(* IEC 61131-3 sources: 2026_Projet_YGO_ExcavatriceDragage/CODE_BACKUP/CODE_20260907_ChantierWeekEnd_v0.6.43/L_SIMULATION, 5 files *)

(* ---- FB_Sim_Encoder.st ---- *)
(* ═══════════════════════════════════════════════════════════════
   🧪 FB_Sim_Encoder — Simulation physique d'un codeur absolu de treuil
   ───────────────────────────────────────────────────────────────
   📄 Doc métier : DOC/AF/AF_Partie-13_Fonction_Simulation_v2.5.md
   🧩 Brique réduite (Partie3 §1bis, "briques E/S & diagnostics") : pas de contrat
      Enable/Reset/Error complet, pas de StartStop/SafeStop — outil de banc, pas
      du métier machine.
   🎯 Rôle : fait "compter" un codeur absolu comme si le treuil tournait
      réellement, à partir des relais de sens commandés et du palier de vitesse courant.
   📥 Enable      : simulation active (SimulationModeActive AND NOT BusEncoderMxIsReal)
   📥 RelayFwd/RelayRev : sens commandé (contacteurs de sens du treuil)
   📥 StepNumber  : palier vitesse courant (1..5) — ex. instWinchM1.StepNumber
      Vitesse = interpolation linéaire : palier 1 → MinSpeedMps (1 m/s), palier 5 → MaxSpeedMps (2 m/s).
   📥 PresetCmd   : TRUE le cycle où un preset (homing) doit être appliqué (PresettTrigCmd = 2)
   📥 PresetValue : valeur brute à charger lors du preset
   📥 SpeedScaleFactor : facteur fin de confort (réglable à chaud, sans recompiler). Défaut 1.0 = vitesse
      réelle telle que définie par MinSpeedMps/MaxSpeedMps/PointsPerRev/CableM_PerRev/CycleTimeS.
   📤 RawPosOut   : position brute simulée (UDINT), à aiguiller à la place de la valeur
      EtherCAT réelle quand le device n'est pas Operational (voir PRG_02_Encoders.st)
   `RawPos` en `VAR_IN_OUT`, référencé depuis `GVL_PERSISTENT`
      (même pattern que `Calib` dans `FB_Encoder_Homing`) — `PERSISTENT` n'est valide que sur du
      `VAR_GLOBAL` en CODESYS, pas sur une variable locale de FB. Un vrai codeur absolu physique
      conserve son comptage brut même à travers un reset FROID (indépendant de l'automate).
   ═══════════════════════════════════════════════════════════════ *)

// === DECLARATION (à coller dans la partie déclaration du POU FB_Sim_Encoder) ===

FUNCTION_BLOCK PUBLIC FB_Sim_Encoder
VAR_INPUT
    Enable           : BOOL;   (* --> [CMD] Active la simulation *)
    RelayFwd         : BOOL;   (* --> [HW] Sens commandé avant *)
    RelayRev         : BOOL;   (* --> [HW] Sens commandé arrière *)
    StepNumber       : INT;    (* --> [CMD] Palier vitesse courant (1..5, 0 = arrêt) *)
    PresetCmd        : BOOL;   (* --> [CMD] Applique un preset (homing) *)
    PresetValue      : UDINT;   (* --> [CFG] Valeur brute à charger au preset *)
    SpeedScaleFactor : REAL := 1.0;   (* --> [CFG] Facteur fin de confort (défaut 1.0) *)
    CoastDistanceM   : REAL := 0.0;   (* --> [CFG] Distance de roulis inertiel apres coupure des relais (m). 0 = arret net (defaut). >0 = le treuil continue a vitesse palier 1 dans le dernier sens sur CoastDistanceM metres -> modelise l'anticipation d'arret mecanique (ex. benne). *)
    PresetLatencyCycles : INT := 3;   (* --> [CFG] Nb cycles automate avant application du preset (referencement non instantane) *)
    TestOffsetCmd    : BOOL;          (* --> [TST] Front montant = applique TestOffsetPts (test banc) *)
    TestOffsetPts    : DINT := 0;     (* --> [TST] Décalage signé à appliquer (points bruts) *)
    // 📐 Paramètres physiques du treuil (mêmes valeurs que FB_Encoder_Scale) + vitesse réelle.
    // Vitesse simulée = interpolation linéaire du palier : palier 1 → MinSpeedMps, palier 5 → MaxSpeedMps.
    MinSpeedMps      : REAL := 1.0;    (* --> [CFG] Vitesse palier 1 (m/s) *)
    MaxSpeedMps      : REAL := 2.0;    (* --> [CFG] Vitesse palier 5 (m/s) *)
    PointsPerRev     : UDINT := 8192;  (* --> [CFG] Résolution codeur (pts/tour) *)
    CableM_PerRev    : REAL := 2.0;    (* --> [CFG] Développement câble (m/tour) *)
    CycleTimeS       : REAL := 0.010;  (* --> [CFG] Période tâche PLC (s) — MainTask 10 ms *)
END_VAR
VAR_OUTPUT
    RawPosOut   : UDINT;   (* <-- [DIAG] Position brute simulée *)
    RawSpdOut   : DINT;    (* <-- [DIAG] Vitesse brute simulée (0x6031:01 en 0.1 RPM) *)
END_VAR
VAR_IN_OUT
    RawPos      : UDINT;   (* <-> [BUS] Référence _SimEncoderRawPosM1/M2 (survit au reset froid) *)
END_VAR
VAR
    Increment      : UDINT;              (* . [LOC] Points ajoutés par cycle *)
    EffStep        : INT;               (* . [LOC] Pas borné (>= 1) *)
    SpeedMps       : REAL;              (* . [LOC] Vitesse simulée (m/s) *)
    TestOffsetEdge : R_TRIG;             (* . [LOC] Front TestOffsetCmd *)
    PresetEdge     : R_TRIG;             (* . [LOC] Front montant PresetCmd *)
    PresetPending  : BOOL;               (* . [LOC] Preset en attente d'application (latence) *)
    PresetCount    : INT;                (* . [LOC] Compteur cycles de latence restants *)
    IncrStep1      : UDINT;              (* . [LOC] Increment par cycle a vitesse palier 1 (pour le roulis) *)
    MovingDir      : INT;                (* . [LOC] Dernier sens actif : +1 avant, -1 arriere, 0 arret *)
    CoastPtsLeft   : REAL;               (* . [LOC] Roulis inertiel restant (points bruts) *)
END_VAR

// === IMPLEMENTATION (à coller dans le corps ST du POU FB_Sim_Encoder) ===

{region "§1 Gate"}
IF NOT Enable THEN
    RawPosOut := RawPos;
    RETURN;
END_IF;
{endregion}

{region "§2 Injection test"}
// Injection test banc : VRAI saut de position (comme un glissement réel),
// pour tester Concept 1 / Méca E ET le rattrapage joystick (voir GVL_Simulation bandeau).
TestOffsetEdge(CLK := TestOffsetCmd);
IF TestOffsetEdge.Q THEN
    RawPos := DINT_TO_UDINT(UDINT_TO_DINT(RawPos) + TestOffsetPts);
END_IF;
{endregion}

{region "§3 Comptage"}
// 🎚️ Vitesse simulée = interpolation linéaire du palier (palier 1 → MinSpeedMps, palier 5 → MaxSpeedMps),
// pas par pas de (Max−Min)/4. Palier 0 (arrêt) ramène au palier 1 mais aucun mouvement n'est
// appliqué tant que RelayFwd/RelayRev = FALSE (section plus bas).
EffStep  := MAX(StepNumber, 1);
SpeedMps := MinSpeedMps + (INT_TO_REAL(EffStep) - 1.0) * ((MaxSpeedMps - MinSpeedMps) / 4.0);
// Points par cycle = vitesse (m/s) × points par mètre × période tâche (s) × facteur confort.
Increment := REAL_TO_UDINT(SpeedMps * (UDINT_TO_REAL(PointsPerRev) / CableM_PerRev) * CycleTimeS * SpeedScaleFactor);
// Increment "lent" (palier 1) : vitesse du roulis inertiel apres coupure des relais.
IncrStep1 := REAL_TO_UDINT(MinSpeedMps * (UDINT_TO_REAL(PointsPerRev) / CableM_PerRev) * CycleTimeS * SpeedScaleFactor);

// Front du preset : lance la latence de referencement (le codeur réel n'est pas
// instantane — il met PresetLatencyCycles cycles a se re-referencer apres le front).
PresetEdge(CLK := PresetCmd);
IF PresetEdge.Q THEN
    PresetPending := TRUE;
    PresetCount := PresetLatencyCycles;
END_IF;

// Pendant l'attente, la position brute est conservee (le codeur n'a pas encore re-reference).
// Le mouvement est gelé pendant la latence, comme un codeur réel en cours de referencement.
IF PresetPending THEN
    IF PresetCount > 0 THEN
        PresetCount := PresetCount - 1;
    ELSE
        // Latence écoulée : applique la valeur cible du preset.
        RawPos := PresetValue;
        PresetPending := FALSE;
    END_IF;
ELSIF RelayFwd THEN
    RawPos := RawPos + Increment;
    MovingDir := 1;
    CoastPtsLeft := CoastDistanceM * (UDINT_TO_REAL(PointsPerRev) / CableM_PerRev);
ELSIF RelayRev THEN
    IF RawPos >= Increment THEN
        RawPos := RawPos - Increment;
    ELSE
        RawPos := 0;
    END_IF;
    MovingDir := -1;
    CoastPtsLeft := CoastDistanceM * (UDINT_TO_REAL(PointsPerRev) / CableM_PerRev);
ELSE
    // Relais coupes : roulis inertiel (anticipation d'arret mecanique). Le treuil
    // continue a vitesse palier 1 dans le dernier sens jusqu'a epuisement de CoastPtsLeft.
    IF (CoastPtsLeft >= 1.0) AND (MovingDir <> 0) THEN
        IF MovingDir = 1 THEN
            RawPos := RawPos + IncrStep1;
        ELSIF RawPos >= IncrStep1 THEN
            RawPos := RawPos - IncrStep1;
        ELSE
            RawPos := 0;
        END_IF;
        CoastPtsLeft := CoastPtsLeft - UDINT_TO_REAL(IncrStep1);
    ELSE
        MovingDir := 0;
        CoastPtsLeft := 0.0;
    END_IF;
END_IF;
{endregion}

{region "§4 Sortie"}
RawPosOut := RawPos;
// Formule inverse vitesse brute EtherCAT CoE (0.1 RPM) :
// SpdValue = (V_mps * 60.0) / (0.1 * CableM_PerRev) = V_mps * 300.0 (sur tambour 2m)
IF (MovingDir <> 0) AND (CableM_PerRev > 0.0) THEN
    IF MovingDir = 1 THEN
        RawSpdOut := REAL_TO_DINT((SpeedMps * 60.0) / (0.1 * CableM_PerRev) * SpeedScaleFactor);
    ELSE
        RawSpdOut := -REAL_TO_DINT((SpeedMps * 60.0) / (0.1 * CableM_PerRev) * SpeedScaleFactor);
    END_IF;
ELSE
    RawSpdOut := 0;
END_IF;
{endregion}

END_FUNCTION_BLOCK

(* ---- FB_Sim_Joystick.st ---- *)
(* ═══════════════════════════════════════════════════════════════
   🧪 FB_Sim_Joystick — Simulation des entrées brutes joystick (bus CAN hors ligne)
   ───────────────────────────────────────────────────────────────
   📄 Doc métier : DOC/AF/AF_Partie-13_Fonction_Simulation_v2.5.md
   🧩 Brique réduite (Partie3 §1bis) : outil de banc, pas du métier machine.
   🎯 Rôle : remplace l'ancien bypass homme-mort codé en dur dans `FB_Joystick`
      (`GVL_DEBUG.DBG_DeadmanBypass_TEST`, qui forçait `DeadmanArmed` en
      permanence — un vrai contournement de sécurité). Ici, on simule les
      ENTRÉES BRUTES du capteur (`RawX`/`RawY`/`RawButton`) : le homme-mort réel
      de `FB_Joystick` reste pleinement actif et doit toujours être "actionné"
      (forcer `RawButton` en instance CODESYS) pour armer — comportement
      métier testé pour de vrai, pas contourné.
   🕹️ Comportement dynamique (conception validée) :
      - Ascending : bouton actif → `RawX`/`RawY` monte de `NeutralRaw` vers la cible
        (0 ou `MaxRaw`) en `RiseTimeS`, avec un bruit pseudo-aléatoire léger.
      - Dépassement (`OvershootActive`) : la cible de montée DÉPASSE la butée
        (MaxRaw+AMT ou 0−AMT) → déclenche le défaut capteur hors plage.
      - Retombée : bouton relâché → descente LINÉAIRE en `FallTimeMs` vers le neutre.
      - Bagotement (`BagotementActive`) : au retour, petit balancement de quelques %
        autour du neutre avant de se stabiliser.
   📥 Enable        : simulation active (SimulationModeActive AND NOT BusJoystickSignalIsReal)
   📥 NeutralRaw    : valeur brute simulée au repos (voir GVL_Simulation.TstJoystickForceNeutralRaw)
   📥 MaxRaw        : valeur brute simulée à fond (voir GVL_Simulation.TstJoystickForceMaxRaw)
   📥 Btn*          : boutons directionnels (1 seul impose une butée d'axe ; 0 ou ≥2 = neutre)
   📥 OvershootActive : bagotement au retour (test mouvement parasite)
   📥 RiseTimeS / FallTimeMs / CycleTimeS : dynamique temporelle (pattern FB_Sim_Encoder)
   📤 RawX/RawY     : valeurs brutes dynamiques (neutre = NeutralRaw)
   📤 RawButton     : homme-mort brut = un bouton directionnel actif
   💡 Note d'application : en vue instance CODESYS, forcer `RawX`/`RawY` à `MaxRaw` (ou une
      valeur intermédiaire) pour simuler un débattement, et `RawButton` à `TRUE` pour simuler
      l'appui homme-mort — exactement comme on forcerait le vrai capteur.
   ═══════════════════════════════════════════════════════════════ *)

// === DECLARATION (à coller dans la partie déclaration du POU FB_Sim_Joystick) ===

FUNCTION_BLOCK PUBLIC FB_Sim_Joystick
VAR_INPUT
    Enable              : BOOL;   (* --> [CMD] Active la simulation *)
    NeutralRaw          : INT := 5000;   (* --> [CFG] Valeur brute au repos (neutre) *)
    MaxRaw              : INT := 10000;   (* --> [CFG] Valeur brute à fond *)
    BtnLeft_Rev_TREMIE  : BOOL;   (* --> [TST] Bouton gauche : X→0, Y→neutre *)
    BtnRight_Fwd_MAINT  : BOOL;   (* --> [TST] Bouton droite : X→MaxRaw, Y→neutre *)
    BtnFwd_Up_Close     : BOOL;   (* --> [TST] Bouton avant : X→neutre, Y→MaxRaw *)
    BtnRev_Down_Open    : BOOL;   (* --> [TST] Bouton arrière : X→neutre, Y→0 *)
    OvershootActive     : BOOL;   (* --> [TST] Dépassement de montée au-delà de 100% (défaut capteur hors plage) *)
    BagotementActive    : BOOL;   (* --> [TST] Bagotement au relâchement (petit balancement autour du neutre) *)
    RiseTimeS           : REAL := 1.5;   (* --> [CFG] Temps de montée 0→100% (s) *)
    FallTimeMs          : TIME := T#200MS;   (* --> [CFG] Temps de retombée 100%→0 *)
    CycleTimeS          : REAL := 0.010;   (* --> [CFG] Période tâche PLC (s) — 10 ms *)
END_VAR
VAR_OUTPUT
    RawX        : INT;   (* <-- [DIAG] Valeur brute axe X (dynamique, neutre = NeutralRaw) *)
    RawY        : INT;   (* <-- [DIAG] Valeur brute axe Y (dynamique, neutre = NeutralRaw) *)
    RawButton   : BOOL;  (* <-- [DIAG] Homme-mort brut = un bouton directionnel actif *)
    ReturningActive : BOOL;  (* <-- [STAT] TRUE si retour dynamique en cours (FALL/OVERSHOOT) — FB_SimBench émet le modèle *)
END_VAR
VAR
    FirstCycle  : BOOL := TRUE;   (* . [LOC] Initialisation au neutre *)
    State       : INT := 0;   (* . [LOC] 0=IDLE, 1=RISE, 2=FALL, 3=OVERSHOOT *)
    TargetX     : INT;   (* . [LOC] Cible brute axe X *)
    TargetY     : INT;   (* . [LOC] Cible brute axe Y *)
    ActiveAxis  : INT;   (* . [LOC] 0=aucun, 1=X, 2=Y (axe en retour) *)
    RiseStep    : REAL;   (* . [LOC] Pas de montée par cycle (points) *)
    FallStep    : REAL;   (* . [LOC] Pas de retombée par cycle (points) *)
    RandCnt     : INT := 0;   (* . [LOC] Compteur pseudo-aléatoire (bruit de montée) *)
    Noise       : INT;   (* . [LOC] Bruit ±25 points (≈ ±0.5% de la course) *)
    BtnCount    : INT;   (* . [LOC] Nombre de boutons directionnels actifs (0..4) *)
    OscDev      : REAL;   (* . [LOC] Écart au neutre de l'oscillateur de bagotement *)
    OscVel      : REAL;   (* . [LOC] Vitesse de l'oscillateur (points/cycle) *)
    OscAcc      : REAL;   (* . [LOC] Accélération de l'oscillateur *)
END_VAR
VAR CONSTANT
    CST_ST_IDLE      : INT := 0;   (* . [CFG] État : au neutre *)
    CST_ST_RISE      : INT := 1;   (* . [CFG] État : montée vers la cible *)
    CST_ST_FALL      : INT := 2;   (* . [CFG] État : retombée linéaire *)
    CST_ST_OVERSHOOT : INT := 3;   (* . [CFG] État : bagotement (oscillations amorties) *)
    CST_OSC_K        : REAL := 0.01;   (* . [CFG] Raideur oscillateur (fréquence bagotement) *)
    CST_OSC_C        : REAL := 0.05;   (* . [CFG] Amortissement (2-3 oscillations visibles) *)
    CST_OVERSHOOT_AMT : INT := 600;   (* . [CFG] Dépassement de montée au-delà de MaxRaw (déclenche défaut capteur hors plage) *)
    CST_BAGOT_AMT     : INT := 500;   (* . [CFG] Amplitude du bagotement au relâchement (~5% autour du neutre) *)
END_VAR

// === IMPLEMENTATION (à coller dans le corps ST du POU FB_Sim_Joystick) ===

{region "§1 Gate"}
// 🔑 Initialise au neutre au premier cycle uniquement ; ensuite RawX/RawY sont pilotés
// dynamiquement par les boutons. Quand la simulation est coupée, on revient au neutre.
IF NOT Enable THEN
    FirstCycle := TRUE;
    State      := CST_ST_IDLE;
    RawX       := NeutralRaw;
    RawY       := NeutralRaw;
    RawButton  := FALSE;
    ReturningActive := FALSE; // 📊 Neutralisation : simulation inactive hors Enable
    RETURN;
END_IF;
{endregion}

{region "§2 Initialisation neutre"}
IF FirstCycle THEN
    RawX       := NeutralRaw;
    RawY       := NeutralRaw;
    RawButton  := FALSE;
    State      := CST_ST_IDLE;
    FirstCycle := FALSE;
END_IF;
{endregion}

{region "§3 Pseudo-aléatoire (bruit de montée)"}
// 🎲 Compteur qui repasse à zéro, multiplié pour rester dans la plage (méthode validée).
// Le bruit s'ajoute à la rampe de montée uniquement (pas à la retombée, linéaire propre).
RandCnt := (RandCnt + 1) MOD 1000;
Noise   := (RandCnt MOD 50) - 25;   // ±25 points (≈ ±0.5% de la course)
{endregion}

{region "§4 Cibles & transitions"}
// 🎯 Un SEUL bouton impose une butée d'axe ; 0 ou ≥2 boutons = neutre (pas de diagonale implicite).
// Si OvershootActive : la cible de montée DÉPASSE la butée (MaxRaw+AMT ou 0−AMT) pour
// déclencher le défaut capteur hors plage (RawOutOfRange) — test du dépassement de valeur.
BtnCount := BOOL_TO_INT(BtnLeft_Rev_TREMIE) + BOOL_TO_INT(BtnRight_Fwd_MAINT)
          + BOOL_TO_INT(BtnFwd_Up_Close) + BOOL_TO_INT(BtnRev_Down_Open);
IF BtnCount = 1 THEN
    IF BtnLeft_Rev_TREMIE THEN
        IF OvershootActive THEN TargetX := 0 - CST_OVERSHOOT_AMT; ELSE TargetX := 0; END_IF;
        TargetY := NeutralRaw; ActiveAxis := 1;
    ELSIF BtnRight_Fwd_MAINT THEN
        IF OvershootActive THEN TargetX := MaxRaw + CST_OVERSHOOT_AMT; ELSE TargetX := MaxRaw; END_IF;
        TargetY := NeutralRaw; ActiveAxis := 1;
    ELSIF BtnFwd_Up_Close THEN
        TargetX := NeutralRaw;
        IF OvershootActive THEN TargetY := MaxRaw + CST_OVERSHOOT_AMT; ELSE TargetY := MaxRaw; END_IF;
        ActiveAxis := 2;
    ELSE
        TargetX := NeutralRaw;
        IF OvershootActive THEN TargetY := 0 - CST_OVERSHOOT_AMT; ELSE TargetY := 0; END_IF;
        ActiveAxis := 2;
    END_IF;
    State := CST_ST_RISE;
ELSE
    // 0 ou ≥2 boutons : retour au neutre.
    TargetX := NeutralRaw;
    TargetY := NeutralRaw;
    IF State = CST_ST_RISE THEN
        // Front de relâchement : retour au neutre. D'abord retombée linéaire (FALL),
        // puis petit bagotement de quelques % autour du neutre si OvershootActive (voir §6).
        State := CST_ST_FALL;
    END_IF;
END_IF;
{endregion}

{region "§5 Ascending (rampe + bruit)"}
IF State = CST_ST_RISE THEN
    // Pas de montée : pleine course (MaxRaw−NeutralRaw) en RiseTimeS.
    RiseStep := INT_TO_REAL(MaxRaw - NeutralRaw) / (RiseTimeS / CycleTimeS);
    // Axe X
    IF RawX < TargetX THEN
        RawX := MIN(RawX + REAL_TO_INT(RiseStep) + Noise, TargetX);
    ELSIF RawX > TargetX THEN
        RawX := MAX(RawX - REAL_TO_INT(RiseStep) - Noise, TargetX);
    END_IF;
    // Axe Y
    IF RawY < TargetY THEN
        RawY := MIN(RawY + REAL_TO_INT(RiseStep) + Noise, TargetY);
    ELSIF RawY > TargetY THEN
        RawY := MAX(RawY - REAL_TO_INT(RiseStep) - Noise, TargetY);
    END_IF;
END_IF;
{endregion}

{region "§6 Retombée linéaire (sans bagotement)"}
IF State = CST_ST_FALL THEN
    // Pas de retombée : pleine course en FallTimeMs (TIME_TO_REAL → ms, /1000 → s).
    FallStep := INT_TO_REAL(MaxRaw - NeutralRaw) / (TIME_TO_REAL(FallTimeMs) / 1000.0 / CycleTimeS);
    IF RawX < NeutralRaw THEN
        RawX := MIN(RawX + REAL_TO_INT(FallStep), NeutralRaw);
    ELSIF RawX > NeutralRaw THEN
        RawX := MAX(RawX - REAL_TO_INT(FallStep), NeutralRaw);
    END_IF;
    IF RawY < NeutralRaw THEN
        RawY := MIN(RawY + REAL_TO_INT(FallStep), NeutralRaw);
    ELSIF RawY > NeutralRaw THEN
        RawY := MAX(RawY - REAL_TO_INT(FallStep), NeutralRaw);
    END_IF;
    IF RawX = NeutralRaw AND RawY = NeutralRaw THEN
        // Arrivée au neutre : si bagotement demandé, lance un petit balancement de quelques %.
        IF BagotementActive THEN
            State := CST_ST_OVERSHOOT;
            IF ActiveAxis = 1 THEN
                OscDev := INT_TO_REAL(CST_BAGOT_AMT);
            ELSE
                OscDev := INT_TO_REAL(CST_BAGOT_AMT);
            END_IF;
            OscVel := 0.0;
        ELSE
            State := CST_ST_IDLE;
        END_IF;
    END_IF;
END_IF;
{endregion}

{region "§7 Bagotement (dépassement + oscillations amorties)"}
IF State = CST_ST_OVERSHOOT THEN
    // 🎢 Oscillateur harmonique amorti discret (semi-implicite) autour du neutre :
    // le joystick dépasse le centre (~12% de l'écart initial) puis oscille 1-2 fois
    // avant de se stabiliser — comportement d'un opérateur qui relâche et balance.
    OscAcc := -CST_OSC_K * OscDev - CST_OSC_C * OscVel;
    OscVel := OscVel + OscAcc;
    OscDev := OscDev + OscVel;
    IF ActiveAxis = 1 THEN
        RawX := NeutralRaw + REAL_TO_INT(OscDev);
    ELSE
        RawY := NeutralRaw + REAL_TO_INT(OscDev);
    END_IF;
    // Stabilisé : revient exactement au centre.
    IF ABS(OscDev) < 1.0 AND ABS(OscVel) < 1.0 THEN
        State := CST_ST_IDLE;
        IF ActiveAxis = 1 THEN
            RawX := NeutralRaw;
        ELSE
            RawY := NeutralRaw;
        END_IF;
    END_IF;
END_IF;
{endregion}

{region "§8 Homme-mort brut + drapeau retour"}
RawButton := BtnLeft_Rev_TREMIE OR BtnRight_Fwd_MAINT OR BtnFwd_Up_Close OR BtnRev_Down_Open;
// Drapeau "retour dynamique en cours" : TRUE si l'état est FALL ou OVERSHOOT (retombée/bagotement).
// Permet à FB_SimBench d'émettre la sortie du modèle même après relâchement du bouton.
ReturningActive := (State = CST_ST_FALL) OR (State = CST_ST_OVERSHOOT);
{endregion}

END_FUNCTION_BLOCK

(* ---- FB_Sim_Safety.st ---- *)
(* ═══════════════════════════════════════════════════════════════
   🧪 FB_Sim_Safety — Simulation de la chaîne d'AU et du contacteur de puissance
   ───────────────────────────────────────────────────────────────
   📥 Enable            : activation de la simulation (SimulationModeActive AND NOT SensorEmergencyStopChainIsReal)
   📥 SimChainOkBit     : bit opérateur — TRUE = simuler la chaîne AU fermée ; FALSE = chaîne ouverte (non simulée)
   📥 PowerCutOff_A     : demande de coupure PLC canal A (TRUE = OK/fermé) — conservé pour interface, non utilisé par SimChainOk
   📥 PowerCutOff_B     : demande de coupure PLC canal B (TRUE = OK/fermé) — conservé pour interface, non utilisé par SimChainOk
   📥 PowerCutOffRequest: requête de coupure métier (PowerCutOffRequest du FB AU) — TRUE = arrêt d'urgence (chaîne ouverte)
   📥 EmergencyArming   : impulsion de réarmement (EmergencyArming_RQ)
   📥 BtnEmergencyStop   : appui coup-de-poing AU (TRUE = boucle ouverte)
   📥 TestCutActive     : test de redondance en cours (canal A ou B coupé par le FB AU)

   📤 SimChainOk        : simulation de la boucle AU (fermée si SimChainOkBit, ouverte sur coup-de-poing/test/coupure)
   📤 SimContactorOk    : simulation du contacteur engagé (PowerContactorEngaged)

   ⚙️ MÉCANISME GRANULAIRE (contrôle opérateur de la chaîne AU) :
      - `SimChainOkBit` pilote la chaîne : FALSE → chaîne OUVERTE (on ne peut pas armer) ;
        TRUE → chaîne FERMÉE (le bouton Armable s'active, on arme, la séquence teste les sorties).
      - Pendant le test de redondance (TestCutActive), la chaîne CLIGNOTE (s'ouvre pendant TEST_A/B,
        se referme pendant RESTORE_A/B) puis revient à 1 — comme en réel.
      - `PowerCutOffRequest` (coupure métier) ouvre la chaîne → ARRÊT D'URGENCE.
      - `BtnEmergencyStop` (coup-de-poing) ouvre la chaîne.
      - Le contacteur ne s'engage QUE pendant l'impulsion d'armement (EmergencyArming), avec une
        temporisation d'engagement (CST_ContactorEngageDelay), puis s'auto-maintient tant que la
        chaîne est saine ; il retombe (CST_ContactorDropDelay) dès que la chaîne s'ouvre.
      - À la ré-entrée en simulation (Enable FALSE→TRUE), SimChainOkBit = FALSE → chaîne OUVERTE et
        contacteur NON engagé (on n'a pas armé) — pas de faux « OK » immédiat.

   🔒 NON-RÉGRESSION ARMEMENT (dépendance circulaire) :
      - La chaîne n'est PAS fermée par défaut : elle est fermée UNIQUEMENT si l'opérateur pose
        `SimChainOkBit`. Elle ne dépend PAS de PowerCutOff_A/B (qui sont dans le cercle) : le
        réarmement après échec de test de redondance (RedundancyTestFailedCause laté → PowerCutOff_A=FALSE)
        reste possible car la chaîne est maintenue fermée par le bit opérateur, pas par le PLC.
      - L'ouverture « PLC coupe un canal » est représentée par TestCutActive (test redondance) et
        PowerCutOffRequest (coupure métier) — jamais par PowerCutOff_A/B seuls.
   ═══════════════════════════════════════════════════════════════
   📄 Doc métier : DOC/AF/AF_Partie-13_Fonction_Simulation_v2.5.md
*)
FUNCTION_BLOCK FB_Sim_Safety
VAR_INPUT
    Enable            : BOOL; // --> [CMD] Activation de la simulation
    SimChainOkBit     : BOOL; // --> [TST] Bit opérateur : TRUE = simuler chaîne AU fermée
    PowerCutOff_A     : BOOL; // --> [SAFE] Commande coupure canal A (TRUE = OK/fermé)
    PowerCutOff_B     : BOOL; // --> [SAFE] Commande coupure canal B (TRUE = OK/fermé)
    PowerCutOffRequest: BOOL; // --> [SAFE] Requête coupure métier (TRUE = arrêt d'urgence)
    EmergencyArming   : BOOL; // --> [CMD] Impulsion de réarmement (TRUE = pulse)
    BtnEmergencyStop   : BOOL; // --> [HW] Force l'ouverture de la boucle (TRUE = bouton appuyé/défaut)
    TestCutActive      : BOOL; // --> [SAFE] Test de redondance en cours (canal A ou B coupé par le FB AU)
END_VAR
VAR_OUTPUT
    SimChainOk      : BOOL; // <-- [STAT] Boucle AU simulée saine
    SimContactorOk  : BOOL; // <-- [STAT] Contacteur simulé engagé
END_VAR
VAR
    ContactorLatch  : BOOL; // . [LOC] Mémorisation de l'auto-maintien du contacteur
    ChainOpenReq    : BOOL; // . [LOC] Demande brute d'ouverture de la chaîne (bit off / coup-de-poing / test / coupure)
    ChainOpen       : BOOL; // . [LOC] État latche de la chaîne (TRUE = ouverte)
    ContactorEngageReq : BOOL; // . [LOC] Demande d'engagement du contacteur (pulse ET chaîne saine)
    TonChainOpen    : TON;  // . [LOC] Temporisation d'ouverture de la chaîne (retombée relais)
    TonChainClose   : TON;  // . [LOC] Temporisation de fermeture de la chaîne (retombée relais)
    TonContactorEngage : TON; // . [LOC] Temporisation d'engagement du contacteur (temps de collage bobine)
    TonContactorDrop   : TON; // . [LOC] Temporisation de retombée du contacteur (temps de décollage bobine)
END_VAR
VAR CONSTANT
    // === TEMPORISATIONS PHYSIQUES SIMULÉES (compatibles séquence FB AU) ===
    // ⚠️ Doivent rester < durées de la séquence FB AU (CST_TestDuration=200ms, CST_ArmingPulseDuration=1s,
    //    CST_ArmingConfirmTimeout=2s) pour que le test de redondance et la confirmation contacteur
    //    restent validés : ouverture/fermeture chaîne < 200ms, engagement contacteur < 1s.
    CST_ChainOpenDelay       : TIME := T#50ms;  // Temps de retombée relais AU (ouverture chaîne)
    CST_ChainCloseDelay      : TIME := T#50ms;  // Temps de retombée relais AU (fermeture chaîne)
    CST_ContactorEngageDelay : TIME := T#100ms; // Temps de collage bobine contacteur (engagement)
    CST_ContactorDropDelay   : TIME := T#50ms;  // Temps de décollage bobine contacteur (retombée)
END_VAR

// === IMPLEMENTATION ===
{region "§1 Gate"}
IF NOT Enable THEN
    SimChainOk     := FALSE;
    SimContactorOk := FALSE;
    ContactorLatch := FALSE;
    ChainOpen      := TRUE; // Chaîne ouverte par défaut à la ré-entrée (on n'a pas armé)
    ChainOpenReq   := FALSE;
    ContactorEngageReq := FALSE;
    TonChainOpen(IN := FALSE);
    TonChainClose(IN := FALSE);
    TonContactorEngage(IN := FALSE);
    TonContactorDrop(IN := FALSE);
    RETURN;
END_IF;
{endregion}

{region "§2 Chaîne AU (contrôle granulaire + dynamique)"}
// 1. La chaîne AU est saine si l'opérateur la simule fermée (SimChainOkBit = TRUE) ET si aucun
//    événement ne l'ouvre : coup-de-poing (BtnEmergencyStop), test de redondance (TestCutActive),
//    coupure métier (PowerCutOffRequest).
// 🔧 DEADLOCK SIMULATION (corrigé) : la chaîne n'est PAS fermée par défaut ni dépendante de
//    PowerCutOff_A/B (qui sont dans le cercle). Elle est fermée UNIQUEMENT par le bit opérateur
//    `SimChainOkBit`. Le réarmement après échec de test de redondance (RedundancyTestFailedCause laté
//    → PowerCutOff_A=FALSE) reste possible car la chaîne est maintenue fermée par le bit, pas par
//    le PLC. Hors simulation (Enable=FALSE), la chaîne reste pilotée par le matériel via le repli
//    HwReal (PRG_02 §1/§2) — aucune régression sécurité réelle.
// 🆕 DYNAMIQUE : l'ouverture/fermeture suit une temporisation (CST_ChainOpenDelay / CST_ChainCloseDelay)
//    qui simule le temps de retombée des relais AU, tout en restant < 200ms (CST_TestDuration) pour
//    ne pas fausser le test de redondance. Pendant le test, la chaîne clignote (s'ouvre en TEST_A/B,
//    se referme en RESTORE_A/B) puis revient à 1.
ChainOpenReq := (NOT SimChainOkBit) OR BtnEmergencyStop OR TestCutActive OR PowerCutOffRequest;

// Temporisation d'ouverture : la chaîne s'ouvre après CST_ChainOpenDelay de demande soutenue
TonChainOpen(IN := ChainOpenReq, PT := CST_ChainOpenDelay);
// Temporisation de fermeture : la chaîne se ferme après CST_ChainCloseDelay d'absence de demande
TonChainClose(IN := NOT ChainOpenReq, PT := CST_ChainCloseDelay);

// Latch de la chaîne avec temporisations (défaut = ouverte à la ré-entrée)
IF ChainOpenReq THEN
    IF TonChainOpen.Q THEN
        ChainOpen := TRUE;
    END_IF;
ELSE
    IF TonChainClose.Q THEN
        ChainOpen := FALSE;
    END_IF;
END_IF;

SimChainOk := NOT ChainOpen;
{endregion}

{region "§3 Auto-maintien contacteur (dynamique réaliste)"}
// 2. Logique d'auto-maintien (latch) du contacteur avec priorité à la coupure.
// 🆕 DYNAMIQUE : le contacteur ne s'engage QUE pendant l'impulsion d'armement (EmergencyArming)
//    tant que la chaîne est saine, après CST_ContactorEngageDelay (temps de collage bobine), puis
//    s'auto-maintient. Il retombe après CST_ContactorDropDelay (temps de décollage bobine) dès que
//    la chaîne s'ouvre — comme une bobine réelle qui décolle sans alimentation. Ces temporisations
//    restent < CST_ArmingPulseDuration (1s) et CST_ArmingConfirmTimeout (2s) pour que la
//    confirmation contacteur reste validée. À la ré-entrée en simulation, le contacteur est NON
//    engagé (on n'a pas armé).
ContactorEngageReq := EmergencyArming AND SimChainOk;

// Temporisation d'engagement : le contacteur se colle après CST_ContactorEngageDelay de pulse soutenu
TonContactorEngage(IN := ContactorEngageReq, PT := CST_ContactorEngageDelay);
// Temporisation de retombée : le contacteur décolle après CST_ContactorDropDelay de chaîne ouverte
TonContactorDrop(IN := NOT SimChainOk, PT := CST_ContactorDropDelay);

// Latch du contacteur avec priorité à la coupure (retombée > engagement)
IF NOT SimChainOk THEN
    IF TonContactorDrop.Q THEN
        ContactorLatch := FALSE;
    END_IF;
ELSIF ContactorEngageReq THEN
    IF TonContactorEngage.Q THEN
        ContactorLatch := TRUE;
    END_IF;
END_IF;

// Recopie vers la sortie
SimContactorOk := ContactorLatch;
{endregion}

(* ---- FB_Sim_Translation.st ---- *)
(* ═══════════════════════════════════════════════════════════════
   🧪 FB_Sim_Translation — Progression capteurs simulés M3
   ───────────────────────────────────────────────────────────────
   🎯 Rôle : Produit les cinq capteurs de position M3 par progression continue
      de Trémie vers Maintenance. Le modèle ne publie que les six mots valides
      de FB_Translation_PositionDecoder : 11111 → 01111 → 00111 → 00011 →
      00001 → 00000.
(* ═══════════════════════════════════════════════════════════════
   🧪 FB_Sim_Translation — Progression capteurs simulés M3
   ───────────────────────────────────────────────────────────────
   🎯 Rôle : Produit les cinq capteurs de position M3 par progression continue
      de Trémie vers Maintenance. Le modèle ne publie que les six mots valides
      de FB_Translation_PositionDecoder : 11111 → 01111 → 00111 → 00011 →
      00001 → 00000.
   📏 Convention : PositionProgress en mètres, 0 m = Trémie … 30 m = Maintenance.
      Distances NON-linéaires : Trémie(0)→PV(5)=5 m, PV(5)→P2(15)=10 m,
      P2(15)→P1(20)=5 m, P1(20)→Maintenance(30)=10 m.
   🔒 Le modèle est une source d'entrée confinée derrière HwIn ; il ne pilote
      aucune sortie réelle. Un override manuel valide est appliqué par
      FB_SimBench, pas par ce FB.
   📄 Doc métier : DOC/AF/AF_Partie-13_Fonction_Simulation_v2.5.md
             DOC/AF/AF_Partie-11_Fonction_Translation_v2.3.md
   ═══════════════════════════════════════════════════════════════ *)

FUNCTION_BLOCK PUBLIC FB_Sim_Translation
VAR_INPUT
    Enable          : BOOL;              (* --> [CMD] TRUE = modèle actif *)
    ReqTremie       : BOOL;              (* --> [CMD] Demande explicite vers Trémie *)
    ReqMaintenance  : BOOL;              (* --> [CMD] Demande explicite vers Maintenance *)
    SpeedTgt_Pct    : REAL;              (* --> [CMD] Magnitude commande 0..100 %, bornée avant calcul *)
    FullTravelTimeS : REAL := 8.0;       (* --> [CFG] Temps complet Trémie→Maintenance à 100 %, simulation seulement *)
END_VAR
VAR_OUTPUT
    PosTremie      : BOOL;               (* <-- [STAT] Bit4 du mot capteurs *)
    PosPV          : BOOL;               (* <-- [STAT] Bit3 du mot capteurs *)
    PosP2          : BOOL;               (* <-- [STAT] Bit2 du mot capteurs (point matériel PVP2) *)
    PosP1          : BOOL;               (* <-- [STAT] Bit1 du mot capteurs *)
    PosMaintenance : BOOL;               (* <-- [STAT] Bit0 du mot capteurs *)
END_VAR
VAR
    instCycleTime              : FB_CycleTime;   (* * [INST] Mesure temps de cycle *)
    PositionProgress           : REAL;   (* . [LOC] 0 m=Trémie ... 30 m=Maintenance *)
    SpeedPctBounded            : REAL;   (* . [LOC] Vitesse bornée *)
    PositionIncrement          : REAL;   (* . [LOC] Incrément de progression *)
    Initialized                : BOOL := FALSE;   (* . [LOC] Initialisation *)
END_VAR
VAR CONSTANT
    // 📏 Positions réelles des 5 capteurs (mètres) — convention 0 m=Trémie, 30 m=Maintenance.
    // Distances NON-linéaires : 0→5 (PV), 5→15 (P2), 15→20 (P1), 20→30 (Maintenance).
    CST_PositionAtTremie       : REAL := 0.0;
    CST_PositionAtPV           : REAL := 5.0;
    CST_PositionAtP2           : REAL := 15.0;
    CST_PositionAtP1           : REAL := 20.0;
    CST_PositionAtMaintenance  : REAL := 30.0;
    CST_TotalDistanceM         : REAL := 30.0; // Distance totale Trémie→Maintenance (m)
    CST_MinFullTravelTimeS     : REAL := 0.1; // Protection division : modèle sans dynamique sous ce seuil
END_VAR

// === IMPLEMENTATION ===

{region "§1 Gate"}
IF NOT Enable THEN
    // Démarrage déterministe au P1 (20 m) = position de travail : mot capteurs 00011
    // (P1 + Maintenance faits). Evite qu'un boot sim en 00000 (tout FALSE) fasse croire
    // au decodeur "extreme Maintenance" et bloque le verrou descente treuil (T249-A).
    PositionProgress := CST_PositionAtP1;
    Initialized := FALSE;
    PosTremie := FALSE;
    PosPV := FALSE;
    PosP2 := FALSE;
    PosP1 := TRUE;
    PosMaintenance := TRUE;
    RETURN;
END_IF;
{endregion}

{region "§2 Initialisation"}
IF NOT Initialized THEN
    PositionProgress := CST_PositionAtP1;   // etat de depart = position de travail P1 (voir §1)
    Initialized := TRUE;
END_IF;
{endregion}

{region "§3 Progression"}
instCycleTime(DefaultValueS := 0.010);
SpeedPctBounded := LIMIT(0.0, ABS(SpeedTgt_Pct), 100.0);

// Une vitesse à 100 % parcourt les 30 m (Trémie→Maintenance) pendant FullTravelTimeS.
// Les demandes de sens sont des bits explicites ; une demande contradictoire est neutre.
IF FullTravelTimeS >= CST_MinFullTravelTimeS THEN
    PositionIncrement := (SpeedPctBounded / 100.0)
                         * (CST_TotalDistanceM / FullTravelTimeS)
                         * instCycleTime.CycleTimeS;
ELSE
    PositionIncrement := 0.0;
END_IF;

IF ReqTremie AND NOT ReqMaintenance THEN
    PositionProgress := MAX(CST_PositionAtTremie, PositionProgress - PositionIncrement);
ELSIF ReqMaintenance AND NOT ReqTremie THEN
    PositionProgress := MIN(CST_PositionAtMaintenance, PositionProgress + PositionIncrement);
END_IF;
{endregion}

{region "§4 Publication capteurs"}
// Réinitialisation explicite : aucune valeur transitoire héritée d'une zone précédente.
PosTremie := FALSE;
PosPV := FALSE;
PosP2 := FALSE;
PosP1 := FALSE;
PosMaintenance := FALSE;

// Chaque intervalle correspond à un seul mot thermomètre valide.
IF PositionProgress <= CST_PositionAtTremie THEN
    PosTremie := TRUE;
    PosPV := TRUE;
    PosP2 := TRUE;
    PosP1 := TRUE;
    PosMaintenance := TRUE;
ELSIF PositionProgress <= CST_PositionAtPV THEN
    PosPV := TRUE;
    PosP2 := TRUE;
    PosP1 := TRUE;
    PosMaintenance := TRUE;
ELSIF PositionProgress <= CST_PositionAtP2 THEN
    PosP2 := TRUE;
    PosP1 := TRUE;
    PosMaintenance := TRUE;
ELSIF PositionProgress <= CST_PositionAtP1 THEN
    PosP1 := TRUE;
    PosMaintenance := TRUE;
ELSIF PositionProgress < CST_PositionAtMaintenance THEN
    PosMaintenance := TRUE;
END_IF;
{endregion}

(* ---- FB_SimBench.st ---- *)
(* ═══════════════════════════════════════════════════════════════
   🧪 FB_SimBench — Enveloppe unique de simulation pour banc d'essai
   ───────────────────────────────────────────────────────────────
   📄 Doc métier : DOC/AF/AF_Partie-13_Fonction_Simulation_v2.5.md

   🎯 Rôle : Compose les 4 blocs de modèle de simulation existants :
      - FB_Sim_Encoder (instM1, instM2)
      - FB_Sim_Translation (instTranslation)
      - FB_Sim_Joystick (instJoystick)
      - FB_Sim_Safety (instSafety)

   🔒 Brique réduite : 0 lecture de variable globale en interne.
      Toutes les entrées (commandes, stimuli, HwReal) sont passées en paramètres.

   🔴 RÈGLES SÉCURITÉ ET POLARITÉ :
      - Modèle frein M1/M2/M3 : M1_BrakeIsOpen_DI := M1_BrakeCmd (1 = OUVERT).
        Ne JAMAIS faire NOT BrakeCmd !
      - Retours contacteurs M1/M2 : 1 = tous retombés (TRUE quand RelayFwd=0 et RelayRev=0).
   ═══════════════════════════════════════════════════════════════ *)

FUNCTION_BLOCK PUBLIC FB_SimBench
VAR_INPUT
    Enable                     : BOOL;             (* --> [CMD] Activation globale (GVL_Simulation.SimulationModeActive) *)

    // ── Commandes issues de l'automate (Scan N-1 / PRG_07 / PRG_10) ──────────
    M1_RelayFwd                : BOOL;   (* --> [CMD] Sens avant M1 *)
    M1_RelayRev                : BOOL;   (* --> [CMD] Sens arrière M1 *)
    // Les 4 contacteurs de palier participent au retour unique
    // « tous contacteurs retombés » — sans eux, le modèle annonce l'arrêt alors qu'un
    // palier est encore engagé (fausse condition d'armement Méca A).
    M1_SpeedContactor_1        : BOOL;   (* --> [HW] Contacteur palier 1 M1 *)
    M1_SpeedContactor_2        : BOOL;   (* --> [HW] Contacteur palier 2 M1 *)
    M1_SpeedContactor_3        : BOOL;   (* --> [HW] Contacteur palier 3 M1 *)
    M1_SpeedContactor_4        : BOOL;   (* --> [HW] Contacteur palier 4 M1 *)
    M1_SpeedCmd_Pct            : REAL;   (* --> [CMD] Consigne vitesse M1 *)
    M1_StepNumber              : INT;    (* --> [CMD] Palier vitesse courant M1 (1..5) *)
    M1_PresetTriggerCmd        : WORD;   (* --> [CMD] Trigger preset M1 *)
    M1_PresetValueOut          : UDINT;   (* --> [CFG] Valeur preset M1 *)
    M1_BrakeCmd                : BOOL;             (* --> [CMD] TRUE = commande desserrage frein M1 *)

    M2_RelayFwd                : BOOL;   (* --> [CMD] Sens avant M2 *)
    M2_RelayRev                : BOOL;   (* --> [CMD] Sens arrière M2 *)
    M2_SpeedContactor_1        : BOOL;   (* --> [HW] Idem M1, voir ci-dessus *)
    M2_SpeedContactor_2        : BOOL;   (* --> [HW] Contacteur palier 2 M2 *)
    M2_SpeedContactor_3        : BOOL;   (* --> [HW] Contacteur palier 3 M2 *)
    M2_SpeedContactor_4        : BOOL;   (* --> [HW] Contacteur palier 4 M2 *)
    M2_SpeedCmd_Pct            : REAL;   (* --> [CMD] Consigne vitesse M2 *)
    M2_StepNumber              : INT;    (* --> [CMD] Palier vitesse courant M2 (1..5) *)
    M2_PresetTriggerCmd        : WORD;   (* --> [CMD] Trigger preset M2 *)
    M2_PresetValueOut          : UDINT;   (* --> [CFG] Valeur preset M2 *)
    M2_BrakeCmd                : BOOL;             (* --> [CMD] TRUE = commande desserrage frein M2 *)

    M3_ReqTremie               : BOOL;             (* --> [CMD] Demande explicite vers Trémie *)
    M3_ReqMaintenance          : BOOL;             (* --> [CMD] Demande explicite vers Maintenance *)
    M3_SpeedCmd_Pct            : REAL;   (* --> [CMD] Consigne vitesse M3 *)
    M3_BrakeCmd                : BOOL;             (* --> [CMD] TRUE = commande desserrage frein M3 *)

    PowerKeepAlive_A           : BOOL;             (* --> [SAFE] TRUE = relais A maintenu sagement par le PLC *)
    PowerKeepAlive_B           : BOOL;             (* --> [SAFE] TRUE = relais B maintenu sagement par le PLC *)
    EmergencyArming_RQ         : BOOL;             (* --> [CMD] Impulsion de réarmement puissance *)
    TestCutActive              : BOOL;             (* --> [SAFE] Test de redondance AU en cours (canal A ou B coupé) *)
    PowerCutOffRequest         : BOOL;             (* --> [SAFE] Requête coupure métier (TRUE = arrêt d'urgence) *)
    SimChainOkBit              : BOOL;             (* --> [TST] Bit opérateur : TRUE = simuler chaîne AU fermée *)

    // ── Stimuli & Paramètres de banc ─────────────────────────────────────────
    SimEncoderSpeedFactor      : REAL := 1.0;   (* --> [CFG] Facteur vitesse codeur *)
    SimWinchCoast_M            : REAL := 0.35;  (* --> [CFG] Roulis inertiel treuils simules apres coupure relais (m) — modelise l'anticipation d'arret meca (benne) ; ~0.35 = finit dans la bande ouvert/ferme malgre l'anticipation d'arret *)
    SimTopPositionActive       : BOOL := FALSE; (* --> [TST] Injection manuelle capteur haut actif (essai ciblé) *)
    SimSyncDeviationInjectM1   : BOOL := FALSE;   (* --> [TST] Injection écart synchro M1 *)
    SimSyncDeviationInjectM2   : BOOL := FALSE;   (* --> [TST] Injection écart synchro M2 *)
    SimSyncDeviationOffset_M   : REAL := 0.5;   (* --> [TST] Offset écart synchro *)

    SimM3SensorsWordOverrideActive : BOOL := FALSE;   (* --> [TST] Override mot capteurs M3 *)
    SimM3SensorsWord               : BYTE := 16#07;   (* --> [TST] Mot capteurs M3 forcé *)

    SimJoystickLeft_Rev_TREMIE_Active  : BOOL := FALSE;   (* --> [TST] Bouton joystick gauche *)
    SimJoystickRight_Fwd_MAINT_Active  : BOOL := FALSE;   (* --> [TST] Bouton joystick droite *)
    SimJoystickFwd_Up_Close_Active     : BOOL := FALSE;   (* --> [TST] Bouton joystick avant *)
    SimJoystickRev_Down_Open_Active    : BOOL := FALSE;   (* --> [TST] Bouton joystick arrière *)
    SimJoystickRawX                    : INT := 5000;   (* --> [TST] Valeur brute X *)
    SimJoystickRawY                    : INT := 5000;   (* --> [TST] Valeur brute Y *)
    SimJoystickRawButton               : BOOL := FALSE;   (* --> [TST] Bouton homme-mort *)
    SimJoystickOvershoot_Active        : BOOL := FALSE;   (* --> [TST] Dépassement de montée au-delà de 100% (défaut capteur hors plage) *)
    SimJoystickBagotement_Active       : BOOL := FALSE;   (* --> [TST] Bagotement au relâchement (petit balancement autour du neutre) *)

    SimKoboldContactValue      : BOOL := FALSE;   (* --> [TST] Contact fond Kobold *)
    BtnEmergencyStop           : BOOL := FALSE;    (* --> [TST] Simulation appui coup-de-poing AU *)

    // ── Image réelle fallback ────────────────────────────────────────────────
    HwReal                     : ST_HardwareImage;   (* --> [HW] Image réelle fallback *)
END_VAR

VAR_OUTPUT
    (* Sorties d'état du profil AF_Partie-03 §2.
       En LD, CODESYS réserve la PREMIÈRE broche de sortie au flux du rung :
       `Ready` n'y porte jamais d'expression, les broches suivantes oui. *)
    Ready                      : BOOL;             (* <-- [STAT] TRUE = banc prêt (Enable actif, modèles à jour) *)
    Busy                       : BOOL;             (* <-- [STAT] TRUE = cycle de simulation en cours *)
    Done                       : BOOL;             (* <-- [STAT] TRUE = images de simulation publiées ce scan *)

    Winch                      : ST_HwWinch;   (* <-- [DIAG] Image treuils simulée *)
    Translation                : ST_HwTranslation;   (* <-- [DIAG] Image translation simulée *)
    Operator                   : ST_HwOperator;   (* <-- [DIAG] Image opérateur simulée *)
    Machine                    : ST_HwMachine;   (* <-- [DIAG] Image machine simulée *)
END_VAR

VAR_IN_OUT
    RawPosM1                   : UDINT;            (* <-> [BUS] Mémoire _SimEncoderRawPosM1 dans GVL_PERSISTENT *)
    RawPosM2                   : UDINT;            (* <-> [BUS] Mémoire _SimEncoderRawPosM2 dans GVL_PERSISTENT *)
END_VAR

VAR CONSTANT
    CST_M3FullTravelTimeS       : REAL := 8.0; // Temps de Trémie à Maintenance à 100 %, modèle banc uniquement
END_VAR

VAR
    // Modèles sous-jacents
    instSimEncoderM1           : FB_Sim_Encoder;   (* * [INST] Modèle codeur M1 *)
    instSimEncoderM2           : FB_Sim_Encoder;   (* * [INST] Modèle codeur M2 *)
    instSimTranslation         : FB_Sim_Translation;   (* * [INST] Modèle translation M3 *)
    instSimJoystick            : FB_Sim_Joystick;   (* * [INST] Modèle joystick *)
    instSimSafety              : FB_Sim_Safety;   (* * [INST] Modèle sécurité *)

    // Calculs internes
    M1_PresetCmd               : BOOL;   (* . [LOC] Trigger preset M1 *)
    M2_PresetCmd               : BOOL;   (* . [LOC] Trigger preset M2 *)
    M1_OffsetPts               : DINT;   (* . [LOC] Offset synchro M1 *)
    M2_OffsetPts               : DINT;   (* . [LOC] Offset synchro M2 *)

    M3_RelayFwd                : BOOL;   (* . [LOC] Sens avant M3 *)
    M3_RelayRev                : BOOL;   (* . [LOC] Sens arrière M3 *)

    SimJoystickDirectionCount  : INT;   (* . [LOC] Nombre de directions actives *)

    M3_ActualFreqHz            : UINT;   (* . [LOC] Fréquence simulée M3 *)
    M3_StatusWordSim           : WORD;   (* . [LOC] StatusWord simulé M3 *)

    // Roulis dynamique avec dispersion pseudo-aléatoire (±0.1m autour de l'anticipation)
    M2_RelayFwdPrev            : BOOL;   (* . [LOC] Mémoire relais Fwd N-1 *)
    M2_RelayRevPrev            : BOOL;   (* . [LOC] Mémoire relais Rev N-1 *)
    RandomSeed                 : UDINT := 123456789; (* . [LOC] Générateur LCG pseudo-aléatoire *)
    M2_EffectiveCoastM         : REAL := 0.35;       (* . [LOC] Distance de roulis M2 courante *)
END_VAR

// === IMPLEMENTATION ===

{region "§1 Repli image reelle banc desactive"}
IF NOT Enable THEN
    // 🔌 Banc désactivé : repli sur l'image réelle, aucune simulation en cours
    Ready       := FALSE;
    Busy        := FALSE;
    Done        := FALSE;
    Winch       := HwReal.Winch;
    Translation := HwReal.Translation;
    Operator    := HwReal.Operator;
    Machine     := HwReal.Machine;
    RETURN;
END_IF;

// ▶️ Banc actif : le cycle de simulation démarre pour ce scan
Ready := TRUE;
Busy  := TRUE;
Done  := FALSE;

{endregion}

{region "§2 Simulation treuils M1/M2"}
// ── 1. MODÈLE TREUILS (M1 + M2) ─────────────────────────────────────────────
// Presets codeurs : déclenchés si PresetTriggerCmd = 2
M1_PresetCmd := (M1_PresetTriggerCmd = 2);
M2_PresetCmd := (M2_PresetTriggerCmd = 2);

// Conversions d'injection d'écart synchro (0.5m -> points codeur avec 8192 pts/tour, 2m/tour)
// 1m = 4096 points codeur.
M1_OffsetPts := REAL_TO_DINT(SimSyncDeviationOffset_M * 4096.0);
M2_OffsetPts := REAL_TO_DINT(SimSyncDeviationOffset_M * 4096.0);

// Instance modèle codeur M1
instSimEncoderM1(
    Enable           := TRUE,
    RelayFwd         := M1_RelayFwd,
    RelayRev         := M1_RelayRev,
    StepNumber       := M1_StepNumber,
    PresetCmd        := M1_PresetCmd,
    PresetValue      := M1_PresetValueOut,
    SpeedScaleFactor := SimEncoderSpeedFactor,
    CoastDistanceM   := SimWinchCoast_M,
    TestOffsetCmd    := SimSyncDeviationInjectM1,
    TestOffsetPts    := M1_OffsetPts,
    RawPos           := RawPosM1
);

// Détection coupure relais M2 pour renouveler la dispersion pseudo-aléatoire (±0.1m)
IF (M2_RelayFwdPrev AND NOT M2_RelayFwd) OR (M2_RelayRevPrev AND NOT M2_RelayRev) THEN
    // Générateur LCG 32-bit standard : X_{n+1} = (1103515245 * X_n + 12345) MOD 2^31
    RandomSeed := (RandomSeed * 1103515245 + 12345) AND 16#7FFFFFFF;
    // Dispersion pseudo-aléatoire entre -0.10 m et +0.10 m
    M2_EffectiveCoastM := SimWinchCoast_M + (UDINT_TO_REAL(RandomSeed MOD 2000) / 10000.0) - 0.10;
END_IF;
M2_RelayFwdPrev := M2_RelayFwd;
M2_RelayRevPrev := M2_RelayRev;

// Instance modèle codeur M2 (avec roulis et dispersion)
instSimEncoderM2(
    Enable           := TRUE,
    RelayFwd         := M2_RelayFwd,
    RelayRev         := M2_RelayRev,
    StepNumber       := M2_StepNumber,
    PresetCmd        := M2_PresetCmd,
    PresetValue      := M2_PresetValueOut,
    SpeedScaleFactor := SimEncoderSpeedFactor,
    CoastDistanceM   := M2_EffectiveCoastM,
    TestOffsetCmd    := SimSyncDeviationInjectM2,
    TestOffsetPts    := M2_OffsetPts,
    RawPos           := RawPosM2
);

// Recopie structures Winch simulées :
// 🛑 POLARITÉ DE FREIN SIMULÉ : 1 = contacteur commandé = frein OUVERT.
// Câblage réel : DI = 1 ⟺ frein OUVERT. Le modèle produit donc M1_BrakeIsOpen_DI := M1_BrakeCmd !
Winch.M1_BrakeIsOpen_DI        := M1_BrakeCmd;
// Retour UNIQUE « tous contacteurs retombés » = sens ET vitesse.
// Omettre les paliers ferait croire à l'arrêt pendant les transitoires → Méca A armée à tort.
Winch.M1_ContactorsReleased_DI := NOT (M1_RelayFwd OR M1_RelayRev
                                    OR M1_SpeedContactor_1 OR M1_SpeedContactor_2
                                    OR M1_SpeedContactor_3 OR M1_SpeedContactor_4);
Winch.M1_ThermalOk_DI          := TRUE; // Sauf panne simulée

Winch.M2_BrakeIsOpen_DI        := M2_BrakeCmd;
Winch.M2_ContactorsReleased_DI := NOT (M2_RelayFwd OR M2_RelayRev
                                    OR M2_SpeedContactor_1 OR M2_SpeedContactor_2
                                    OR M2_SpeedContactor_3 OR M2_SpeedContactor_4);
Winch.M2_ThermalOk_DI          := TRUE;

// Cohérent avec M2_TensionedCable_DI (sain par défaut) : capteur TOP libre en simu,
// sauf stimulus manuel SimTopPositionActive (injection de fait capteur au banc).
Winch.M1M2_TopPositionFree_DI  := NOT SimTopPositionActive;
Winch.M2_TensionedCable_DI     := TRUE; // Câble tendu en simu

Winch.COD1_PosValue            := instSimEncoderM1.RawPosOut;
Winch.COD1_SpdValue            := instSimEncoderM1.RawSpdOut;
Winch.COD1_Alarms              := 0;
Winch.COD1_Warnings            := 0;
Winch.COD1_DeviceState         := DEVICE_STATE.RUNNING; // État device RUNNING (bus OK)

Winch.COD2_PosValue            := instSimEncoderM2.RawPosOut;
Winch.COD2_SpdValue            := instSimEncoderM2.RawSpdOut;
Winch.COD2_Alarms              := 0;
Winch.COD2_Warnings            := 0;
Winch.COD2_DeviceState         := DEVICE_STATE.RUNNING; // État device RUNNING

{endregion}

{region "§3 Simulation translation M3"}
// ── 2. MODÈLE TRANSLATION M3 (AC600) ─────────────────────────────────────────
M3_RelayFwd := M3_ReqTremie AND NOT M3_ReqMaintenance;
M3_RelayRev := M3_ReqMaintenance AND NOT M3_ReqTremie;

instSimTranslation(
    Enable          := TRUE,
    ReqTremie       := M3_RelayFwd,
    ReqMaintenance  := M3_RelayRev,
    SpeedTgt_Pct    := M3_SpeedCmd_Pct,
    FullTravelTimeS := CST_M3FullTravelTimeS
);

// Remplissage capteurs de position M3 : l'override manuel conserve exactement le
// même ordre que FB_Translation_PositionDecoder (bit4=Trémie ... bit0=Maintenance).
IF SimM3SensorsWordOverrideActive THEN
    Translation.M3_PosTremie_DI      := SimM3SensorsWord.4;
    Translation.M3_PosPV_DI          := SimM3SensorsWord.3;
    Translation.M3_PosPVP2_DI        := SimM3SensorsWord.2;
    Translation.M3_PosP1_DI          := SimM3SensorsWord.1;
    Translation.M3_PosMaintenance_DI := SimM3SensorsWord.0;
ELSE
    Translation.M3_PosTremie_DI      := instSimTranslation.PosTremie;
    Translation.M3_PosPV_DI          := instSimTranslation.PosPV;
    Translation.M3_PosPVP2_DI        := instSimTranslation.PosP2;
    Translation.M3_PosP1_DI          := instSimTranslation.PosP1;
    Translation.M3_PosMaintenance_DI := instSimTranslation.PosMaintenance;
END_IF;

// Polarité frein M3 (1 = OUVERT)
Translation.M3_BrakeIsOpen_DI    := M3_BrakeCmd;

// Thermique moteur/variateur AC600 — pas de panne simulée, toujours OK (comme Winch.M1/M2_ThermalOk_DI)
Translation.M3_ThermalOK_DI      := TRUE;

// Simulation StatusWord AC600 : Bit 0 (Power Ready) = 1, Bit 7 (Comm Ready) = 1 -> 16#0087 en mouvement
// Bit0 retombe à l'arrêt, cohérent avec un variateur qui confirme l'arrêt sans rester "actif" —
// FB_Safety_Translation lit ce bit comme indicateur "mouvement non commandé" (Méca B, TonMecaB 3s) :
// un Bit0 forcé à 1 en continu à l'arrêt déclencherait un PowerCutOff simulé permanent après 3s.
// DrivePowerReady (diagnostic IHM seul, non consommé par un interlock) est le seul autre lecteur,
// aucune régression de mouvement possible.
IF M3_RelayFwd OR M3_RelayRev THEN
    M3_StatusWordSim := 16#0087; // + Operating/Running
    M3_ActualFreqHz  := REAL_TO_UINT(M3_SpeedCmd_Pct * 50.0); // 50.0 Hz à 100% (x100 -> 5000)
ELSE
    M3_StatusWordSim := 16#0080; // Comm Ready seul -- Bit0 retombé, arrêt confirmé
    M3_ActualFreqHz  := 0;
END_IF;

Translation.M3_StatusWord        := M3_StatusWordSim;
Translation.M3_ActualFrequencyHz := M3_ActualFreqHz;
Translation.AC600_DeviceState    := DEVICE_STATE.RUNNING; // État device RUNNING

{endregion}

{region "§4 Simulation operateur joystick"}
// ── 3. MODÈLE OPÉRATEUR / JOYSTICK ───────────────────────────────────────────
instSimJoystick(
    Enable              := TRUE,
    NeutralRaw          := 5000,
    MaxRaw              := 10000,
    BtnLeft_Rev_TREMIE  := SimJoystickLeft_Rev_TREMIE_Active,
    BtnRight_Fwd_MAINT  := SimJoystickRight_Fwd_MAINT_Active,
    BtnFwd_Up_Close     := SimJoystickFwd_Up_Close_Active,
    BtnRev_Down_Open    := SimJoystickRev_Down_Open_Active,
    OvershootActive     := SimJoystickOvershoot_Active,
    BagotementActive    := SimJoystickBagotement_Active,
    CycleTimeS          := 0.010
);

// Les boutons directionnels simplifient les essais : une commande unique impose
// une butée d'axe ; aucune commande ou une combinaison reste au neutre / stimulus avancé.
// Le modèle dynamique (montée/retombée/bagotement) pilote RawX/RawY dès qu'un bouton est actif.
SimJoystickDirectionCount := BOOL_TO_INT(SimJoystickLeft_Rev_TREMIE_Active)
                           + BOOL_TO_INT(SimJoystickRight_Fwd_MAINT_Active)
                           + BOOL_TO_INT(SimJoystickFwd_Up_Close_Active)
                           + BOOL_TO_INT(SimJoystickRev_Down_Open_Active);
IF (SimJoystickDirectionCount >= 1) OR instSimJoystick.ReturningActive THEN
    // Bouton(s) actif(s) OU retour dynamique en cours (retombée/bagotement) → sortie du modèle.
    // (≥2 boutons : le modèle gère lui-même le neutre — pas de diagonale implicite.)
    Operator.JoyXRaw_ANA1 := instSimJoystick.RawX;
    Operator.JoyYRaw_ANA2 := instSimJoystick.RawY;
ELSE
    // Modèle au repos → stimulus analogique avancé (mode « sans bouton »).
    Operator.JoyXRaw_ANA1 := SimJoystickRawX;
    Operator.JoyYRaw_ANA2 := SimJoystickRawY;
END_IF;

// Homme-mort : stimulus brut amont. En simulation avec boutons directionnels actifs,
// l'appui homme-mort est automatiquement inclus pour faciliter les essais sur banc.
Operator.JoyBtnRaw := SimJoystickRawButton OR (SimJoystickDirectionCount > 0);

Operator.CanBusState      := 2; // CANbusState 2 = ACTIVE
Operator.JOY1_DeviceState := DEVICE_STATE.RUNNING; // État device RUNNING

{endregion}

{region "§5 Simulation securite et image machine"}
// ── 4. MODÈLE SÉCURITÉ & COMMUNS MACHINE ─────────────────────────────────────
instSimSafety(
    Enable            := TRUE,
    SimChainOkBit     := SimChainOkBit,
    PowerCutOff_A     := PowerKeepAlive_A,
    PowerCutOff_B     := PowerKeepAlive_B,
    PowerCutOffRequest:= PowerCutOffRequest,
    EmergencyArming   := EmergencyArming_RQ,
    BtnEmergencyStop  := BtnEmergencyStop,
    TestCutActive     := TestCutActive
);

Machine.PowerContactorEngaged_DI   := instSimSafety.SimContactorOk;
Machine.EmergencyChainClosed_DI    := instSimSafety.SimChainOk;
Machine.PhaseRotationOk_DI             := TRUE;
Machine.M1_M2_M3_BrakeThermalOk_DI     := TRUE;
Machine.M1_M2_KoboldBottomTouch_DI     := SimKoboldContactValue;
Machine.HydraulicThermalOk_DI          := TRUE;
Machine.TremieFull_OR_GateRaised_DI    := FALSE; // Pas encore câblé, simulé inactif par défaut

// ✅ Cycle de simulation terminé : les 4 images sont publiées pour ce scan
Busy := FALSE;
Done := TRUE;

{endregion}

END_FUNCTION_BLOCK
